{attribute 'qualified_only'}
{attribute 'strict'}
TYPE E_CIP_Client_Selector :
(
	eNone := 0,
	eClose,
	eFuture,
	eMarinade_Up,
	eMarinade_Low,
	eColor_Up,
	eColor_Low,
	eDrain,
	eLoop
);
END_TYPE

(* stored: Version 1.1.0.1, ProductVersion 3.1.4024.12
   DUT E_CIP_Client_Selector: Id {7051611e-ea40-40c5-adb3-e4b44481b3a3} *)
